// SIMATIC S7-200 project (STEP 7-Micro/WIN), CPU 224XP CN REL 02.01

SYMBOL_TABLE USUARIO1
SO               I0.3
S_I              I0.4
SM               I0.5
S1               I0.7
S2               I1.0
S3               I1.1
SBB1             I1.3
SBB2             I1.2
QS               I1.4
SA               I1.5
am               Q0.0
C_1              Q0.4
C_2              Q0.5
C_3              Q0.6
HL1              Q0.7
HL2              Q1.0
HL3              Q1.1
E0               M0.0
E1               M0.1
E2               M0.2
E3               M0.3
E4               M0.4
E5               M0.5
E6               M0.6
E7               M0.7
E8               M1.0
E9               M1.1
E10              M1.2
E11              M1.3
E12              M1.4
E13              M1.5
E14              M1.6
EM               M1.7
MOTOR            M2.0
E15              M2.1
E16              M2.2
END_SYMBOL_TABLE

ORGANIZATION_BLOCK PRINCIPAL:OB1
TITLE=UNIDAD DE SELECCION
BEGIN
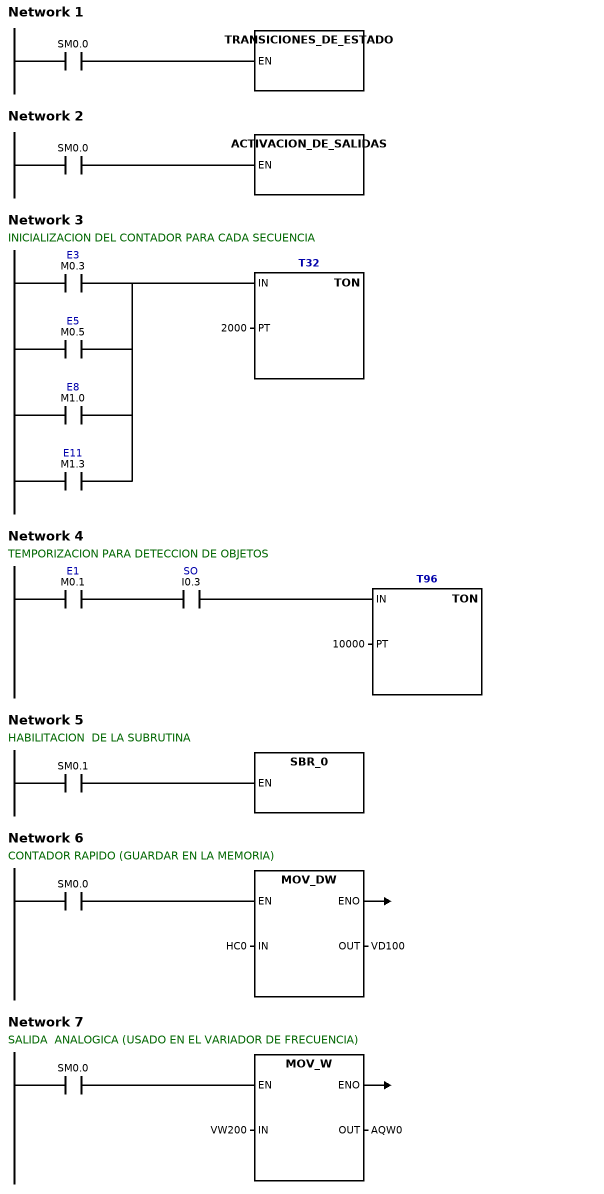
Network 1
LD     SM0.0
CALL   TRANSICIONES_DE_ESTADO:SBR1
Network 2
LD     SM0.0
CALL   ACTIVACION_DE_SALIDAS:SBR2
Network 3
// INICIALIZACION DEL CONTADOR PARA CADA SECUENCIA 
LD     E3:M0.3
O      E5:M0.5
O      E8:M1.0
O      E11:M1.3
TON    T32, 2000
Network 4
// TEMPORIZACION PARA DETECCION DE OBJETOS
LD     E1:M0.1
A      SO:I0.3
TON    T96, 10000
Network 5
// HABILITACION  DE LA SUBRUTINA
LD     SM0.1
CALL   SBR_0:SBR0
Network 6
// CONTADOR RAPIDO (GUARDAR EN LA MEMORIA)
LD     SM0.0
MOVD   HC0, VD100
Network 7
// SALIDA  ANALOGICA (USADO EN EL VARIADOR DE FRECUENCIA)
LD     SM0.0
MOVW   VW200, AQW0
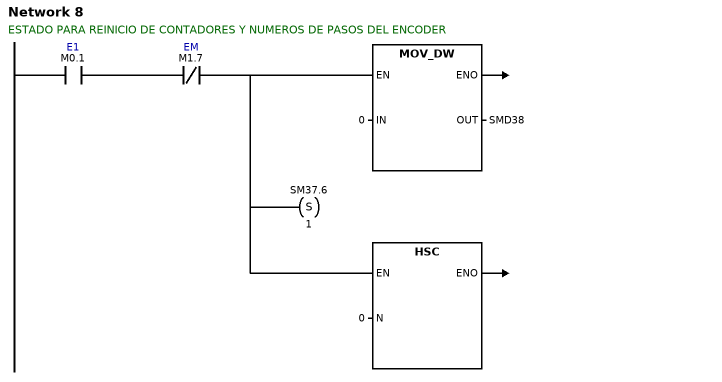
Network 8
// ESTADO PARA REINICIO DE CONTADORES Y NUMEROS DE PASOS DEL ENCODER
LD     E1:M0.1
AN     EM:M1.7
MOVD   0, SMD38
S      SM37.6, 1
HSC    0
END_ORGANIZATION_BLOCK

SUBROUTINE_BLOCK SBR_0:SBR0
TITLE=COMENTARIOS DE LA SUBRUTINA
BEGIN
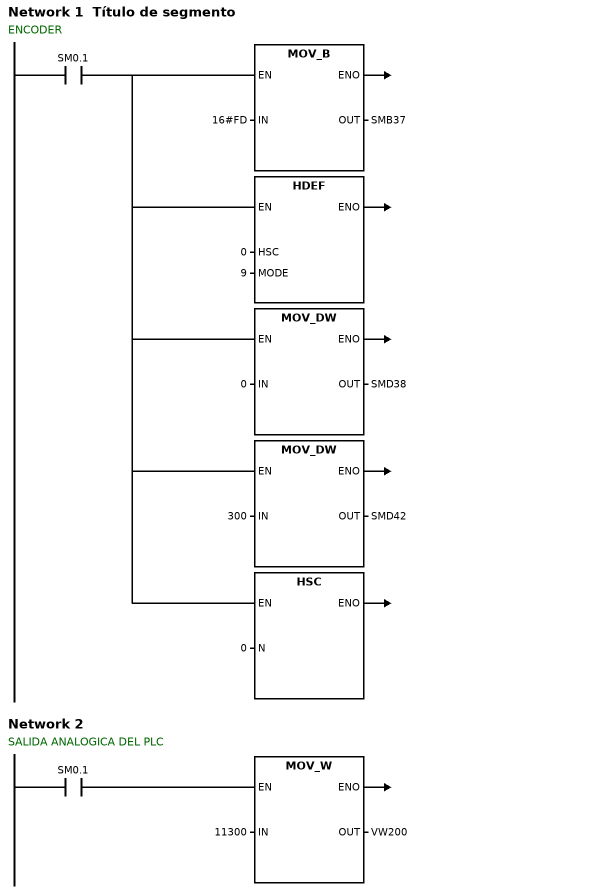
Network 1 // Título de segmento
// ENCODER
LD     SM0.1
MOVB   16#FD, SMB37
HDEF   0, 9
MOVD   0, SMD38
MOVD   300, SMD42
HSC    0
Network 2
// SALIDA ANALOGICA DEL PLC 
LD     SM0.1
MOVW   11300, VW200
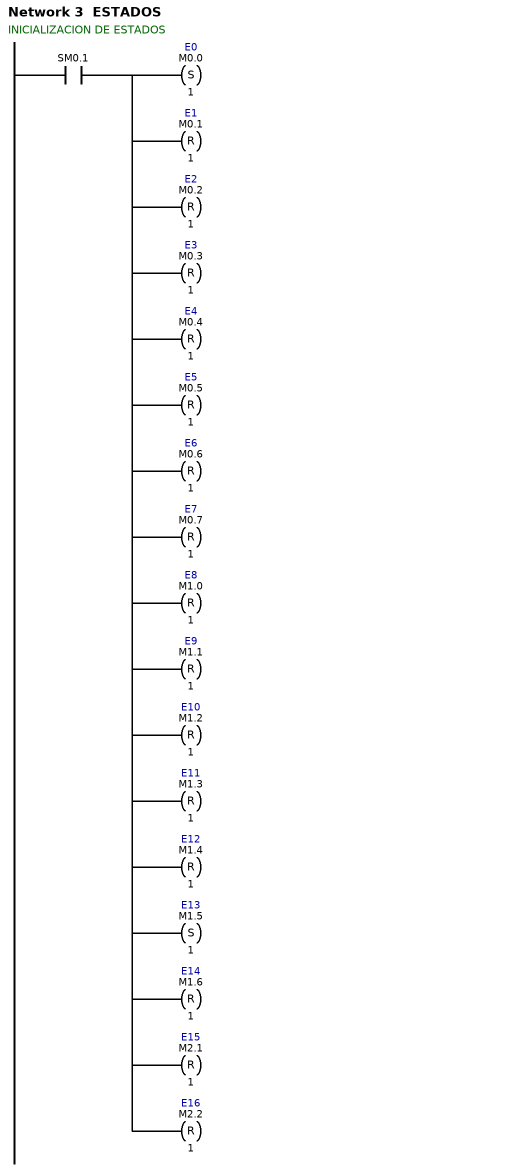
Network 3 // ESTADOS
// INICIALIZACION DE ESTADOS
LD     SM0.1
S      E0:M0.0, 1
R      E1:M0.1, 1
R      E2:M0.2, 1
R      E3:M0.3, 1
R      E4:M0.4, 1
R      E5:M0.5, 1
R      E6:M0.6, 1
R      E7:M0.7, 1
R      E8:M1.0, 1
R      E9:M1.1, 1
R      E10:M1.2, 1
R      E11:M1.3, 1
R      E12:M1.4, 1
S      E13:M1.5, 1
R      E14:M1.6, 1
R      E15:M2.1, 1
R      E16:M2.2, 1
Network 4 // INICIALIZACION DE ESTADOS
END_SUBROUTINE_BLOCK

SUBROUTINE_BLOCK TRANSICIONES_DE_ESTADO:SBR1
TITLE=TRANSICIONES DE ESTADO
BEGIN
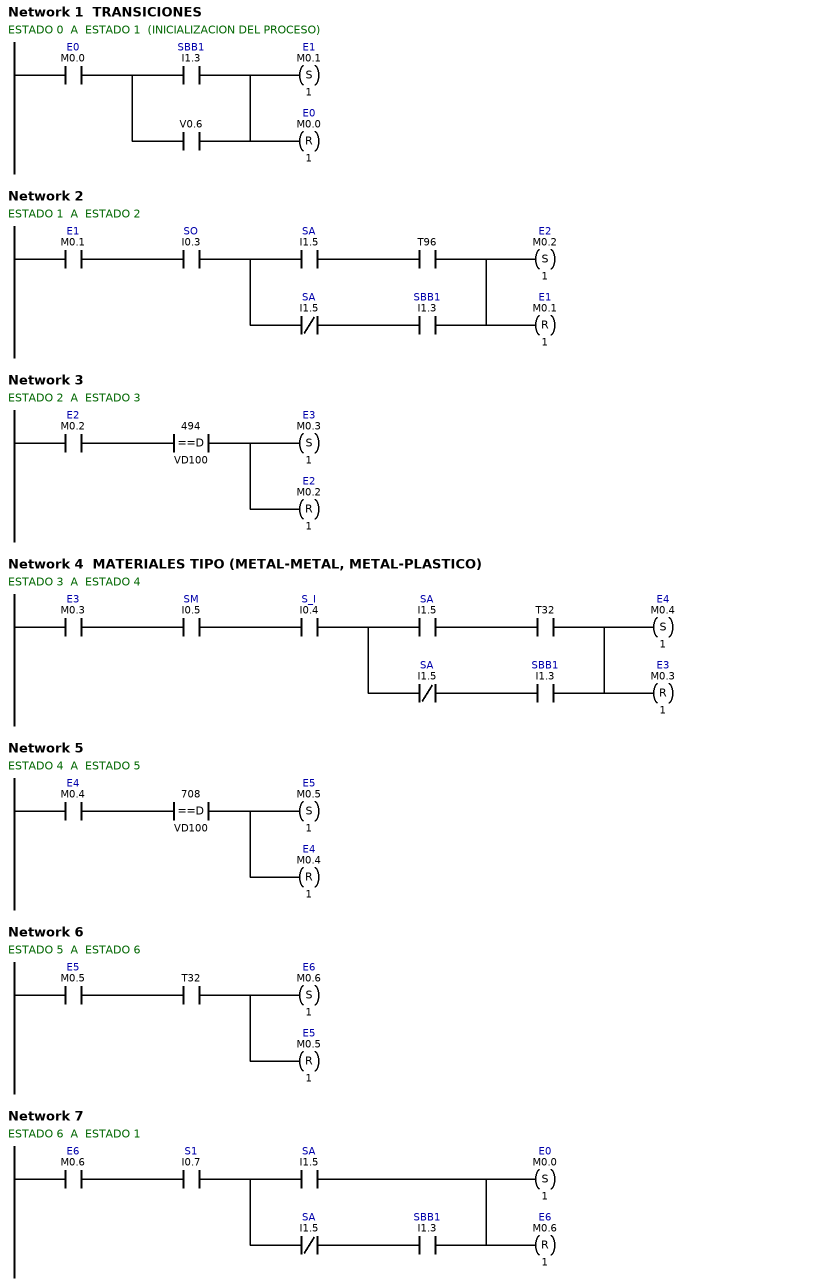
Network 1 // TRANSICIONES
// ESTADO 0  A  ESTADO 1  (INICIALIZACION DEL PROCESO)
LD     E0:M0.0
LD     SBB1:I1.3
O      V0.6
ALD
S      E1:M0.1, 1
R      E0:M0.0, 1
Network 2
// ESTADO 1  A  ESTADO 2 
LD     E1:M0.1
A      SO:I0.3
LD     SA:I1.5
A      T96
LDN    SA:I1.5
A      SBB1:I1.3
OLD
ALD
S      E2:M0.2, 1
R      E1:M0.1, 1
Network 3
// ESTADO 2  A  ESTADO 3
LD     E2:M0.2
AD=    494, VD100
S      E3:M0.3, 1
R      E2:M0.2, 1
Network 4 // MATERIALES TIPO (METAL-METAL, METAL-PLASTICO)
// ESTADO 3  A  ESTADO 4
LD     E3:M0.3
A      SM:I0.5
A      S_I:I0.4
LD     SA:I1.5
A      T32
LDN    SA:I1.5
A      SBB1:I1.3
OLD
ALD
S      E4:M0.4, 1
R      E3:M0.3, 1
Network 5
// ESTADO 4  A  ESTADO 5
LD     E4:M0.4
AD=    708, VD100
S      E5:M0.5, 1
R      E4:M0.4, 1
Network 6
// ESTADO 5  A  ESTADO 6
LD     E5:M0.5
A      T32
S      E6:M0.6, 1
R      E5:M0.5, 1
Network 7
// ESTADO 6  A  ESTADO 1
LD     E6:M0.6
A      S1:I0.7
LD     SA:I1.5
LDN    SA:I1.5
A      SBB1:I1.3
OLD
ALD
S      E0:M0.0, 1
R      E6:M0.6, 1
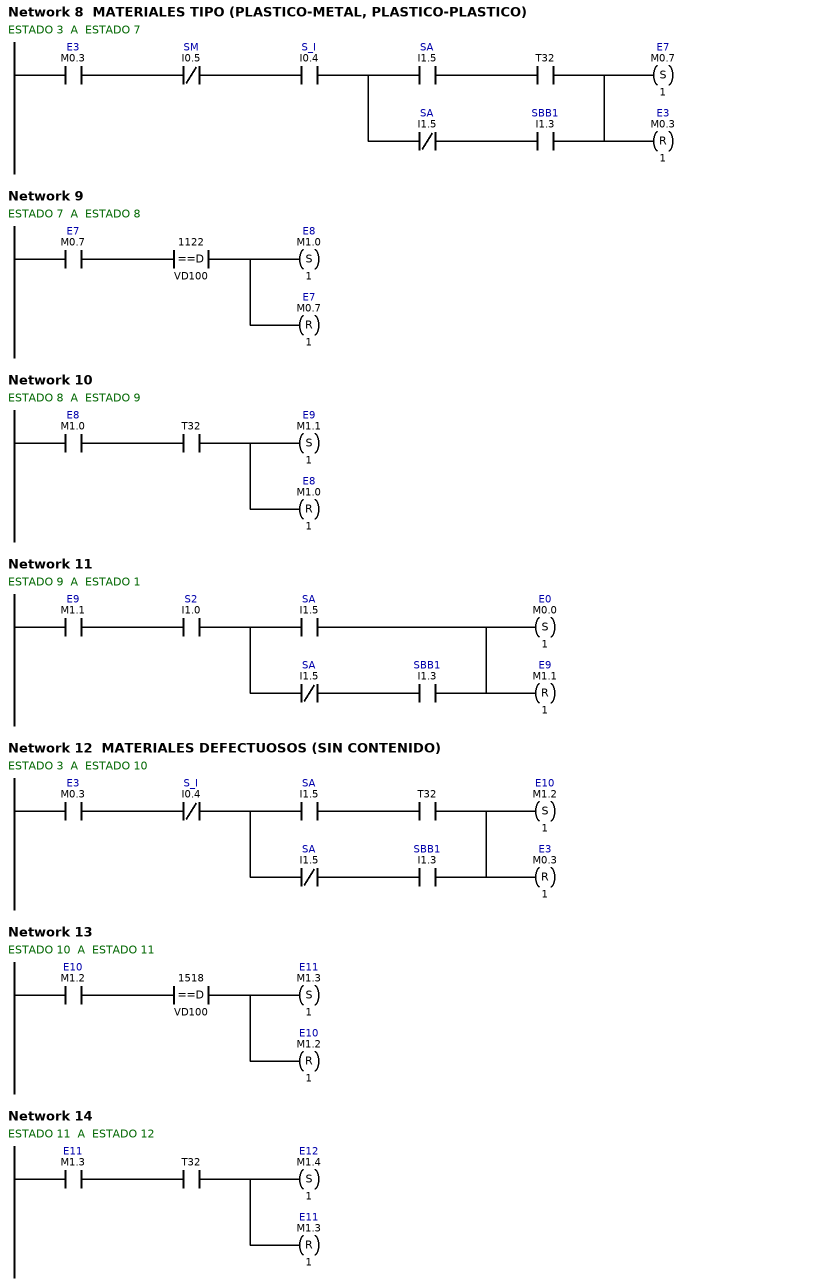
Network 8 // MATERIALES TIPO (PLASTICO-METAL, PLASTICO-PLASTICO)
// ESTADO 3  A  ESTADO 7
LD     E3:M0.3
AN     SM:I0.5
A      S_I:I0.4
LD     SA:I1.5
A      T32
LDN    SA:I1.5
A      SBB1:I1.3
OLD
ALD
S      E7:M0.7, 1
R      E3:M0.3, 1
Network 9
// ESTADO 7  A  ESTADO 8
LD     E7:M0.7
AD=    1122, VD100
S      E8:M1.0, 1
R      E7:M0.7, 1
Network 10
// ESTADO 8  A  ESTADO 9
LD     E8:M1.0
A      T32
S      E9:M1.1, 1
R      E8:M1.0, 1
Network 11
// ESTADO 9  A  ESTADO 1
LD     E9:M1.1
A      S2:I1.0
LD     SA:I1.5
LDN    SA:I1.5
A      SBB1:I1.3
OLD
ALD
S      E0:M0.0, 1
R      E9:M1.1, 1
Network 12 // MATERIALES DEFECTUOSOS (SIN CONTENIDO)
// ESTADO 3  A  ESTADO 10 
LD     E3:M0.3
AN     S_I:I0.4
LD     SA:I1.5
A      T32
LDN    SA:I1.5
A      SBB1:I1.3
OLD
ALD
S      E10:M1.2, 1
R      E3:M0.3, 1
Network 13
// ESTADO 10  A  ESTADO 11
LD     E10:M1.2
AD=    1518, VD100
S      E11:M1.3, 1
R      E10:M1.2, 1
Network 14
// ESTADO 11  A  ESTADO 12
LD     E11:M1.3
A      T32
S      E12:M1.4, 1
R      E11:M1.3, 1
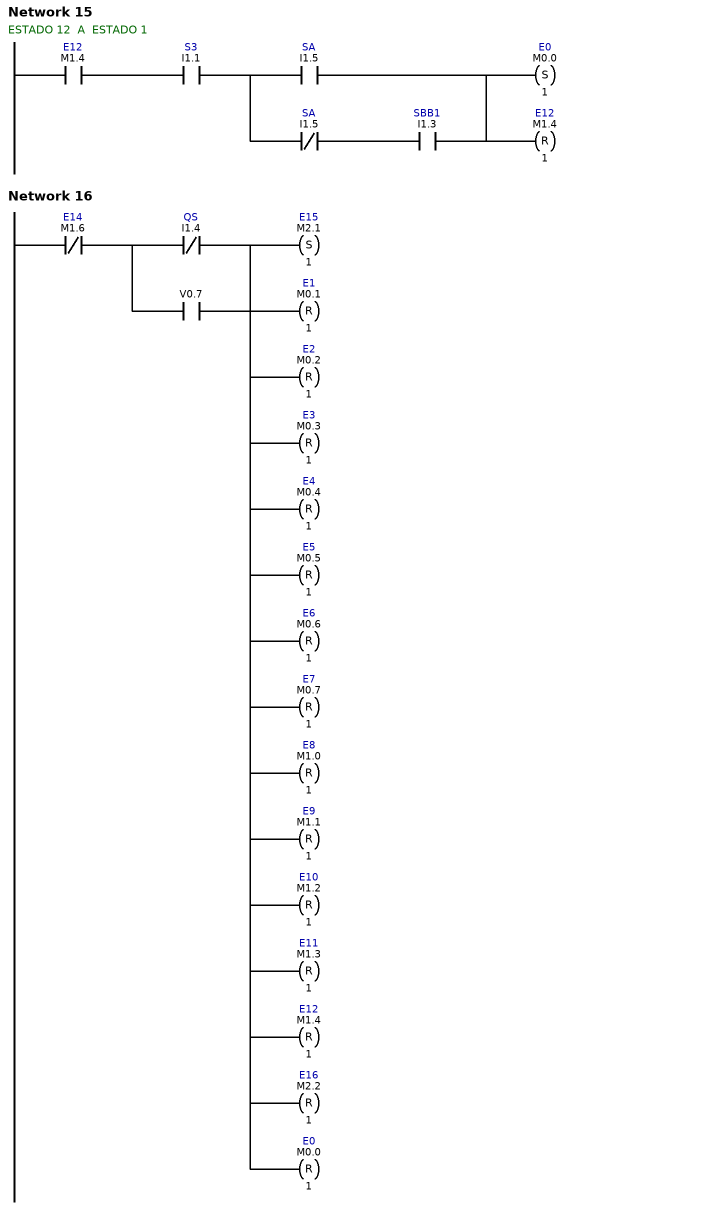
Network 15
// ESTADO 12  A  ESTADO 1
LD     E12:M1.4
A      S3:I1.1
LD     SA:I1.5
LDN    SA:I1.5
A      SBB1:I1.3
OLD
ALD
S      E0:M0.0, 1
R      E12:M1.4, 1
Network 16
// (network saved uncompiled; LAD cells follow)
// row 0: c0 -|/|- E14:M1.6 v  c1 -|/|- QS:I1.4 v  c2 -(S) E15:M2.1, 1
// row 1: c0 ^  c1 -| |- V0.7 ^v  c2 -(R) E1:M0.1, 1
// row 2: c1 ^v  c2 -(R) E2:M0.2, 1
// row 3: c1 ^v  c2 -(R) E3:M0.3, 1
// row 4: c1 ^v  c2 -(R) E4:M0.4, 1
// row 5: c1 ^v  c2 -(R) E5:M0.5, 1
// row 6: c1 ^v  c2 -(R) E6:M0.6, 1
// row 7: c1 ^v  c2 -(R) E7:M0.7, 1
// row 8: c1 ^v  c2 -(R) E8:M1.0, 1
// row 9: c1 ^v  c2 -(R) E9:M1.1, 1
// row 10: c1 ^v  c2 -(R) E10:M1.2, 1
// row 11: c1 ^v  c2 -(R) E11:M1.3, 1
// row 12: c1 ^v  c2 -(R) E12:M1.4, 1
// row 13: c1 ^v  c2 -(R) E16:M2.2, 1
// row 14: c1 ^  c2 -(R) E0:M0.0, 1
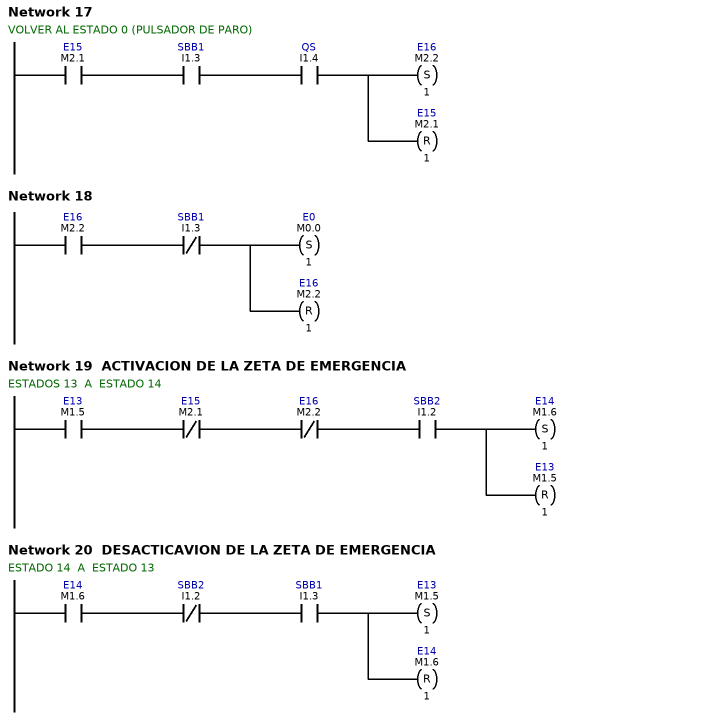
Network 17
// VOLVER AL ESTADO 0 (PULSADOR DE PARO)
LD     E15:M2.1
A      SBB1:I1.3
A      QS:I1.4
S      E16:M2.2, 1
R      E15:M2.1, 1
Network 18
LD     E16:M2.2
AN     SBB1:I1.3
S      E0:M0.0, 1
R      E16:M2.2, 1
Network 19 // ACTIVACION DE LA ZETA DE EMERGENCIA
// ESTADOS 13  A  ESTADO 14
LD     E13:M1.5
AN     E15:M2.1
AN     E16:M2.2
A      SBB2:I1.2
S      E14:M1.6, 1
R      E13:M1.5, 1
Network 20 // DESACTICAVION DE LA ZETA DE EMERGENCIA
// ESTADO 14  A  ESTADO 13
LD     E14:M1.6
AN     SBB2:I1.2
A      SBB1:I1.3
S      E13:M1.5, 1
R      E14:M1.6, 1
Network 21 // Título de segmento
// Comentario de segmento
END_SUBROUTINE_BLOCK

SUBROUTINE_BLOCK ACTIVACION_DE_SALIDAS:SBR2
TITLE=COMENTARIOS DE LA SUBRUTINA
BEGIN
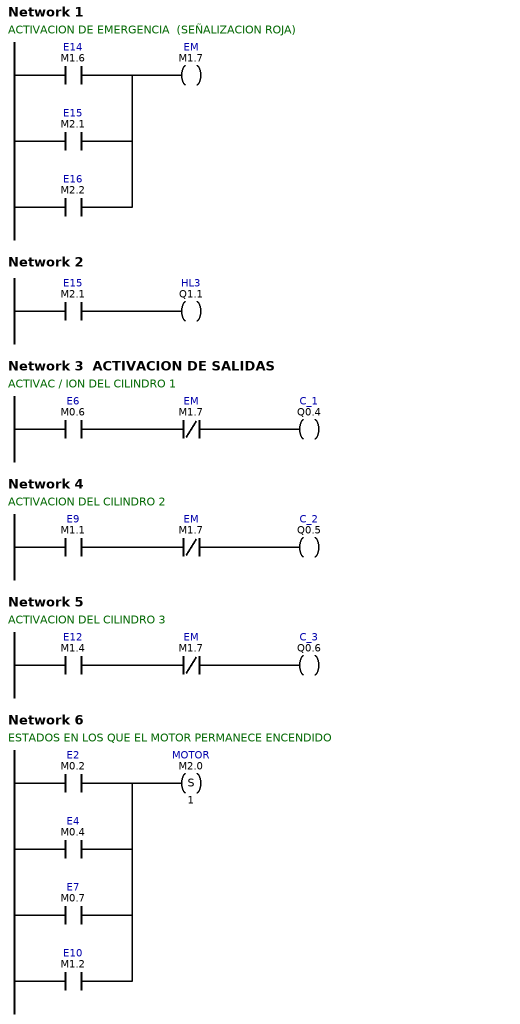
Network 1
// ACTIVACION DE EMERGENCIA  (SEÑALIZACION ROJA)
LD     E14:M1.6
O      E15:M2.1
O      E16:M2.2
=      EM:M1.7
Network 2
LD     E15:M2.1
=      HL3:Q1.1
Network 3 // ACTIVACION DE SALIDAS
// ACTIVAC
// ION DEL CILINDRO 1
LD     E6:M0.6
AN     EM:M1.7
=      C_1:Q0.4
Network 4
// ACTIVACION DEL CILINDRO 2
LD     E9:M1.1
AN     EM:M1.7
=      C_2:Q0.5
Network 5
// ACTIVACION DEL CILINDRO 3
LD     E12:M1.4
AN     EM:M1.7
=      C_3:Q0.6
Network 6
// ESTADOS EN LOS QUE EL MOTOR PERMANECE ENCENDIDO
LD     E2:M0.2
O      E4:M0.4
O      E7:M0.7
O      E10:M1.2
S      MOTOR:M2.0, 1
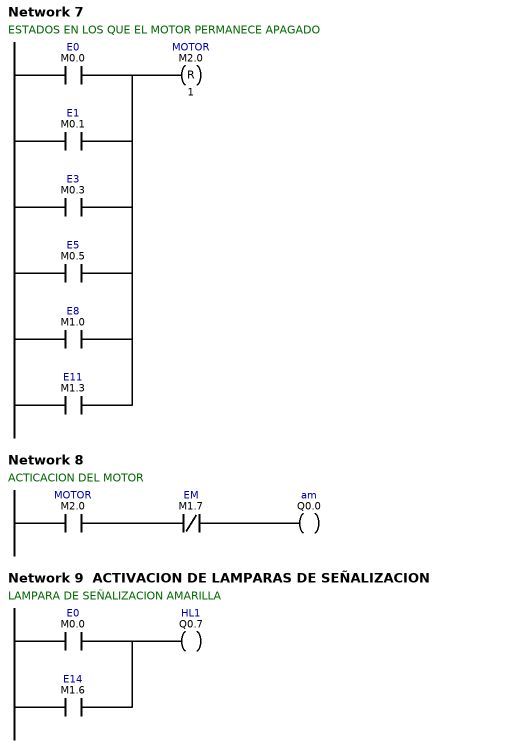
Network 7
// ESTADOS EN LOS QUE EL MOTOR PERMANECE APAGADO
LD     E0:M0.0
O      E1:M0.1
O      E3:M0.3
O      E5:M0.5
O      E8:M1.0
O      E11:M1.3
R      MOTOR:M2.0, 1
Network 8
// ACTICACION DEL MOTOR
LD     MOTOR:M2.0
AN     EM:M1.7
=      am:Q0.0
Network 9 // ACTIVACION DE LAMPARAS DE SEÑALIZACION
// LAMPARA DE SEÑALIZACION AMARILLA
LD     E0:M0.0
O      E14:M1.6
=      HL1:Q0.7
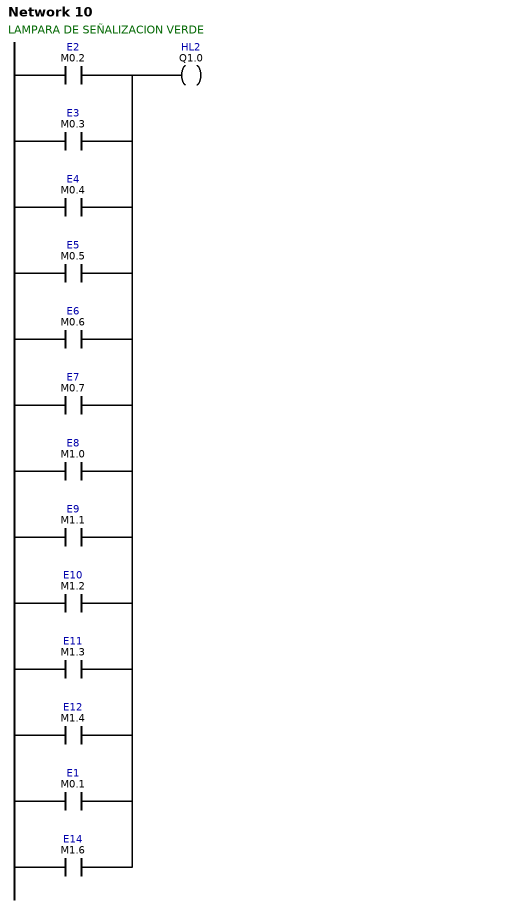
Network 10
// LAMPARA DE SEÑALIZACION VERDE
LD     E2:M0.2
O      E3:M0.3
O      E4:M0.4
O      E5:M0.5
O      E6:M0.6
O      E7:M0.7
O      E8:M1.0
O      E9:M1.1
O      E10:M1.2
O      E11:M1.3
O      E12:M1.4
O      E1:M0.1
O      E14:M1.6
=      HL2:Q1.0
Network 11 // Título de segmento
// Comentario de segmento
END_SUBROUTINE_BLOCK
